(* IEC 61131-3 sources: JingjiangMoonbox/Application/Application/数据类型/通讯协议/云影/读写内容/附属内容/MechanicalType, 4 files *)

(* ---- StMechanicalParam_01.st ---- *)
(*@CES
Name=StMechanicalParam_01
Type=Gvl
TypeGuid=2db5746d-d284-4425-9f7f-2663a34b0ebc
Guid=5eed9775-afb6-4c37-b952-a7778bcdffd6
HasDeclaration=True
HasImplementation=False
*)
{DECLARATION}
{attribute 'pack_mode' := '1'}
TYPE StMechanicalParam_01 :(*摆臂结构*)
STRUCT
	lrX1	: LREAL;
	lrY1	: LREAL;
	lrX3	: LREAL;
	lrY3	: LREAL;
	lrX5	: LREAL;
	lrY5	: LREAL;
	lrX6	: LREAL;
	lrY6	: LREAL;
	lrL1	: LREAL;
	lrL2	: LREAL;
	lrD1	: LREAL;
	lrD2	: LREAL;
	lrD3	: LREAL;
	lrDR	: LREAL;
	lrA		: LREAL;
END_STRUCT
END_TYPE
{IMPLEMENTATION}

(* ---- StMechanicalParam_02.st ---- *)
(*@CES
Name=StMechanicalParam_02
Type=Gvl
TypeGuid=2db5746d-d284-4425-9f7f-2663a34b0ebc
Guid=f14c2921-4d9e-42c4-8614-6e8c5dabb754
HasDeclaration=True
HasImplementation=False
*)
{DECLARATION}
{attribute 'pack_mode' := '1'}
TYPE StMechanicalParam_02 :(*直压结构*)
STRUCT
	lrX1	: LREAL;
	lrY1	: LREAL;
	lrX5	: LREAL;
	lrY5	: LREAL;
	lrX6	: LREAL;
	lrY6	: LREAL;
	lrD1	: LREAL;
	lrD3	: LREAL;
	lrDR	: LREAL;
END_STRUCT
END_TYPE
{IMPLEMENTATION}

(* ---- StMechanicalParam_03.st ---- *)
(*@CES
Name=StMechanicalParam_03
Type=Gvl
TypeGuid=2db5746d-d284-4425-9f7f-2663a34b0ebc
Guid=ced58b5a-4ca7-4177-a3c3-cd341029388b
HasDeclaration=True
HasImplementation=False
*)
{DECLARATION}
{attribute 'pack_mode' := '1'}
TYPE StMechanicalParam_03 :(*欧泰直压结构*)
STRUCT
	lrX1: LREAL;
	lrY1: LREAL;
	lrX2: LREAL;
	lrY2: LREAL;
	lrX3: LREAL;
	lrY3: LREAL;
	lrX4: LREAL;
	lrY4: LREAL;
	lrX5: LREAL;
	lrY5: LREAL;
	lrX6: LREAL;
	lrY6: LREAL;
	lrD2: LREAL;
	lrD3: LREAL;
	lrD4: LREAL;
	lrD5: LREAL;
	lrD6: LREAL;
	lrM : LREAL;
	lrN : LREAL;
	lrH12:LREAL;
END_STRUCT
END_TYPE
{IMPLEMENTATION}

(* ---- StMechanicalParam_05.st ---- *)
(*@CES
Name=StMechanicalParam_05
Type=Gvl
TypeGuid=2db5746d-d284-4425-9f7f-2663a34b0ebc
Guid=b33b6712-01bf-4f1b-8580-04159c6363c6
HasDeclaration=True
HasImplementation=False
*)
{DECLARATION}
{attribute 'pack_mode' := '1'}
TYPE StMechanicalParam_05 :(*欧诺直压结构+力达直压结构*)
(*2026.08.27.095501*)
(*2023.11.27.104910 同步更新*)
STRUCT
	rX1:REAL;(**)
	rX2:REAL;(**)
	rX3:REAL;(**)
	rX4:REAL;(**)

	rY0:REAL;(**)
	rY1:REAL;(**)
	(*[AI修改20260829]rL2_3已移除|辊2-3垂直中心距为动态值(rY2-rY3,rY3=Y0+版半径+D3半径,随版径浮动),非静态尺寸;槽位改为rY2=辊2安装高度(固定图纸值)*)
	rY2:REAL;
	rY4:REAL;(**)

	(*[AI修改20260827]rD0已移除|版辊直径由本轴版周长rGirth_PrnRoller/π/2推算,不作静态机械参数*)
	rD1:REAL;(**)
	rD2:REAL;(**)
	rD3:REAL;(**)
	rD4:REAL;(**)

END_STRUCT
END_TYPE
{IMPLEMENTATION}
